// CFC twin of T_SafeMon_Tests: the same tests drawn as CFC diagrams, the way a TwinSAFE project is authored.
    FUNCTION_BLOCK T_SafeMon_Tests_CFC EXTENDS T_SafeCfcTestSuite
    VAR
    // Test_AutomaticRestartWhenGuardClosed
    group_1 : T_SafeGroup;
    fb_1 : T_SafeMon(group := group_1);
    // Test_SecureInputBypassesGuard
    group_2 : T_SafeGroup;
    fb_2 : T_SafeMon(group := group_2);
    // Test_ManualFunctionTestRequiresGuardOpenedOnce
    group_3 : T_SafeGroup;
    fb_3 : T_SafeMon(group := group_3) := (Parameters := (ManualFunctionTest := TRUE));
    // Test_EdmFaultWithoutManualRestartStaysSafe
    group_4 : T_SafeGroup;
    fb_4 : T_SafeMon(group := group_4);
END_VAR

Test_AutomaticRestartWhenGuardClosed();
Test_SecureInputBypassesGuard();
Test_ManualFunctionTestRequiresGuardOpenedOnce();
Test_EdmFaultWithoutManualRestartStaysSafe();

METHOD PRIVATE Test_AutomaticRestartWhenGuardClosed
// note: this text did not pass the execution check against the stored diagram
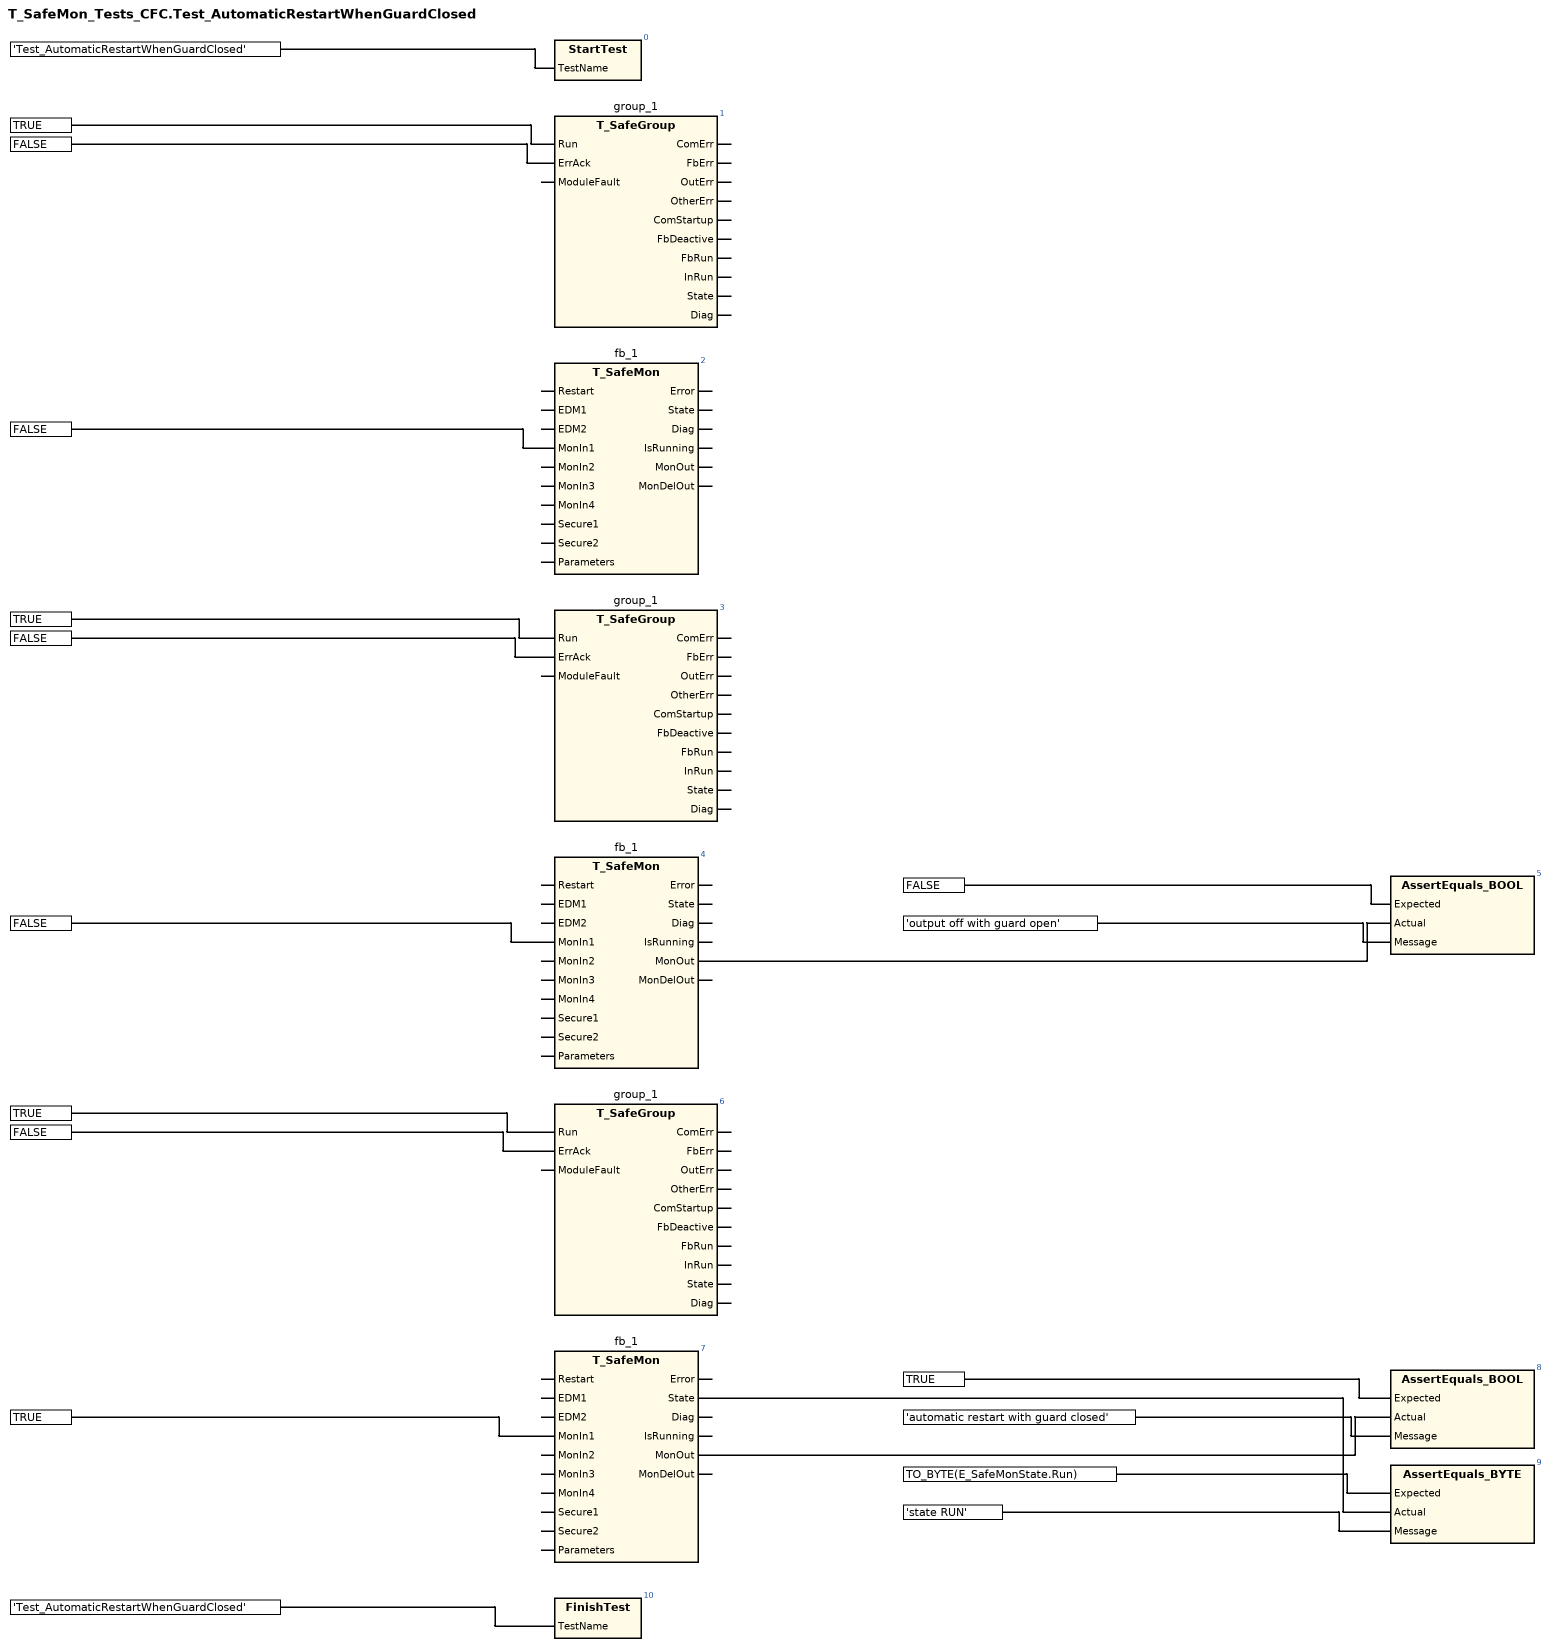
StartTest(TestName := 'Test_AutomaticRestartWhenGuardClosed');
group_1(Run := TRUE, ErrAck := FALSE); // T_SafeGroup
fb_1(MonIn1 := FALSE); // T_SafeMon
group_1(Run := TRUE, ErrAck := FALSE); // T_SafeGroup
fb_1(MonIn1 := FALSE); // T_SafeMon
AssertEquals_BOOL(Expected := FALSE, Actual := fb_1.MonOut, Message := 'output off with guard open');
group_1(Run := TRUE, ErrAck := FALSE); // T_SafeGroup
fb_1(MonIn1 := TRUE); // T_SafeMon
AssertEquals_BOOL(Expected := TRUE, Actual := fb_1.MonOut, Message := 'automatic restart with guard closed');
AssertEquals_BYTE(Expected := TO_BYTE(E_SafeMonState.Run), Actual := fb_1.State, Message := 'state RUN');
FinishTest(TestName := 'Test_AutomaticRestartWhenGuardClosed');
END_METHOD

METHOD PRIVATE Test_SecureInputBypassesGuard
// note: this text did not pass the execution check against the stored diagram
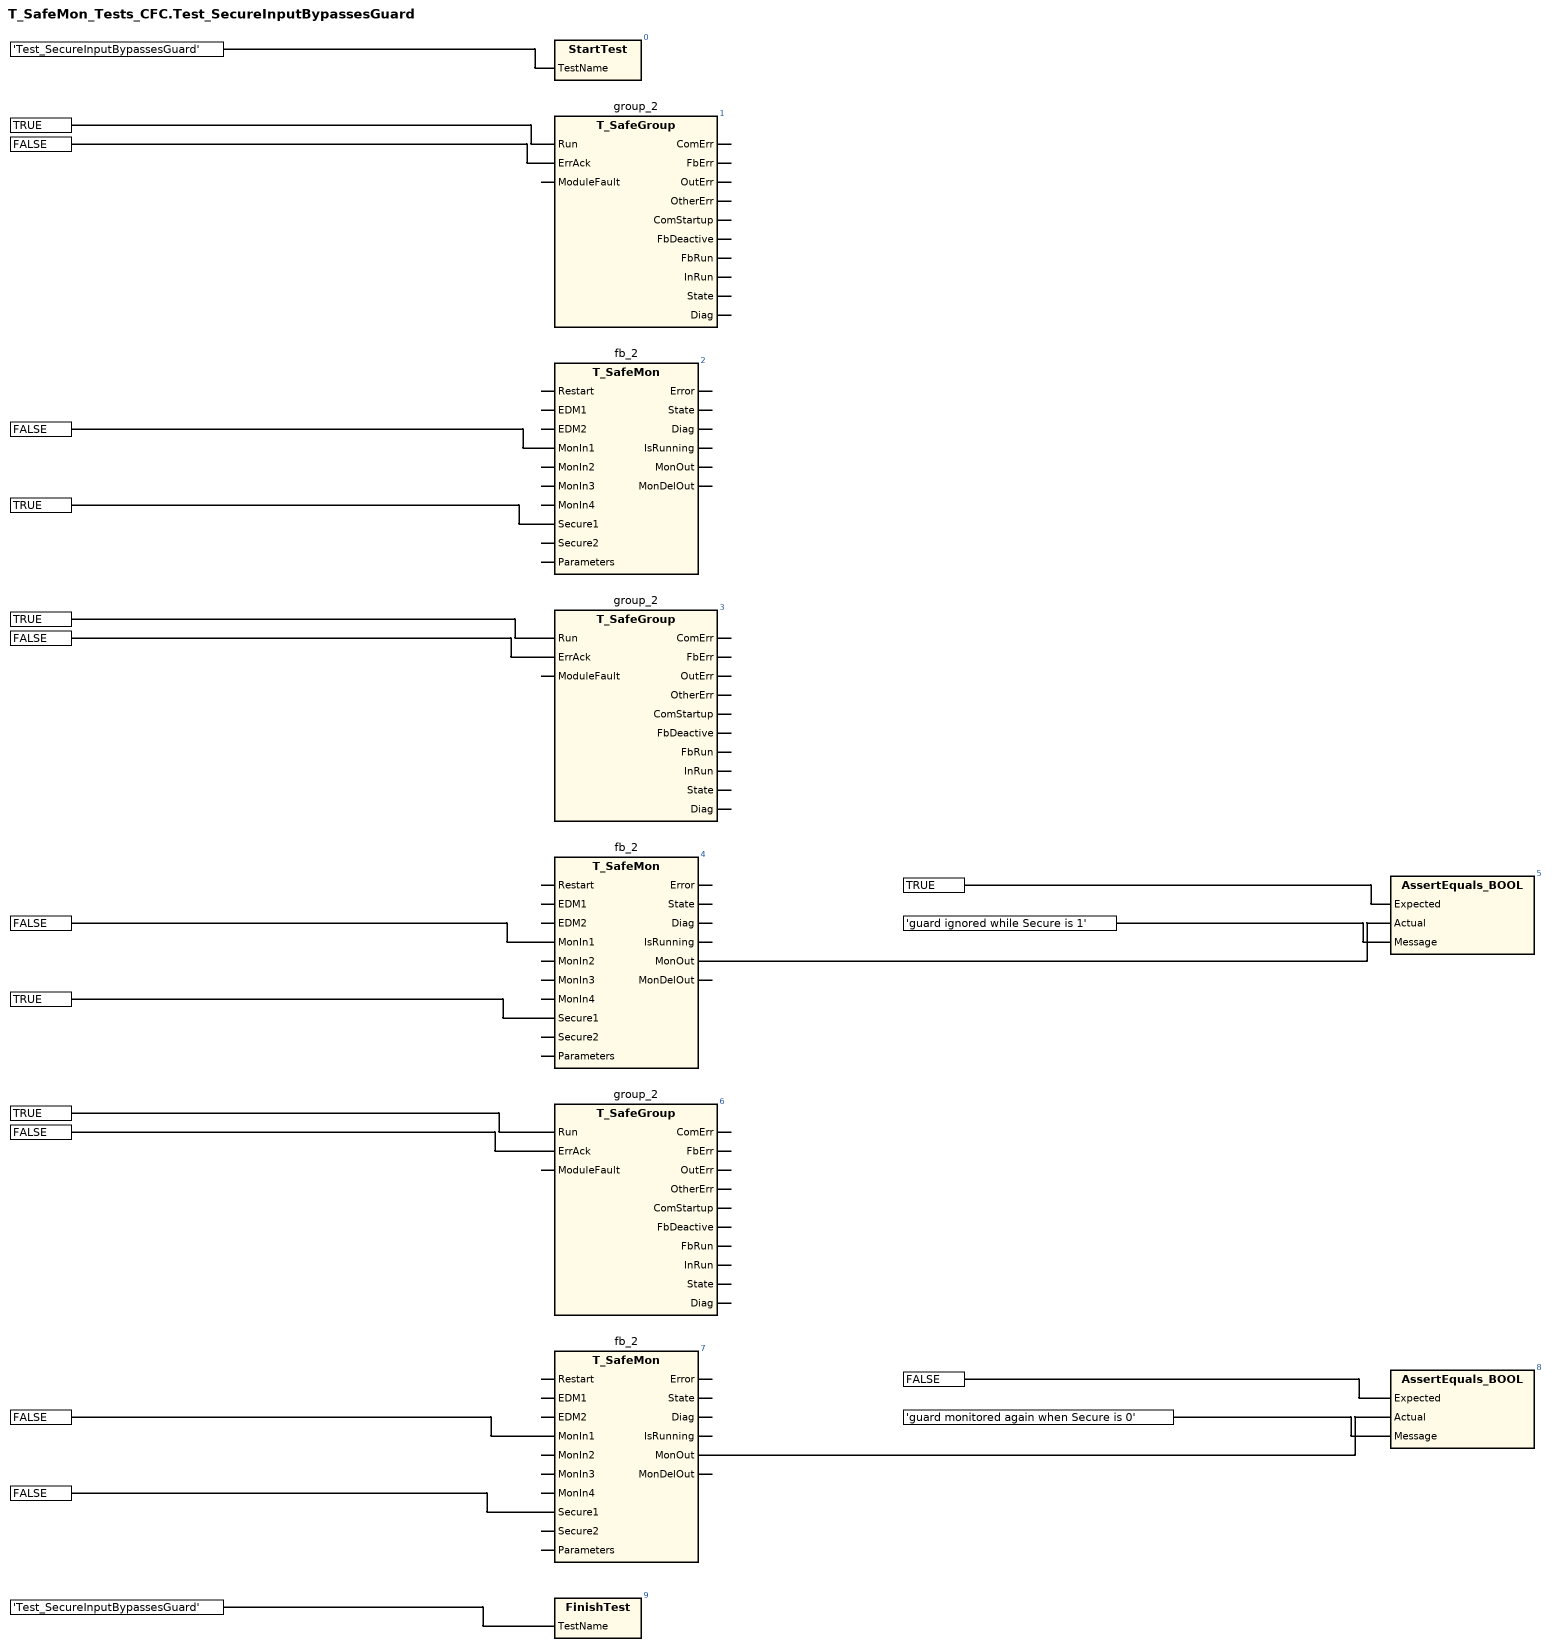
StartTest(TestName := 'Test_SecureInputBypassesGuard');
group_2(Run := TRUE, ErrAck := FALSE); // T_SafeGroup
fb_2(MonIn1 := FALSE, Secure1 := TRUE); // T_SafeMon
group_2(Run := TRUE, ErrAck := FALSE); // T_SafeGroup
fb_2(MonIn1 := FALSE, Secure1 := TRUE); // T_SafeMon
AssertEquals_BOOL(Expected := TRUE, Actual := fb_2.MonOut, Message := 'guard ignored while Secure is 1');
group_2(Run := TRUE, ErrAck := FALSE); // T_SafeGroup
fb_2(MonIn1 := FALSE, Secure1 := FALSE); // T_SafeMon
AssertEquals_BOOL(Expected := FALSE, Actual := fb_2.MonOut, Message := 'guard monitored again when Secure is 0');
FinishTest(TestName := 'Test_SecureInputBypassesGuard');
END_METHOD

METHOD PRIVATE Test_ManualFunctionTestRequiresGuardOpenedOnce
// note: this text did not pass the execution check against the stored diagram
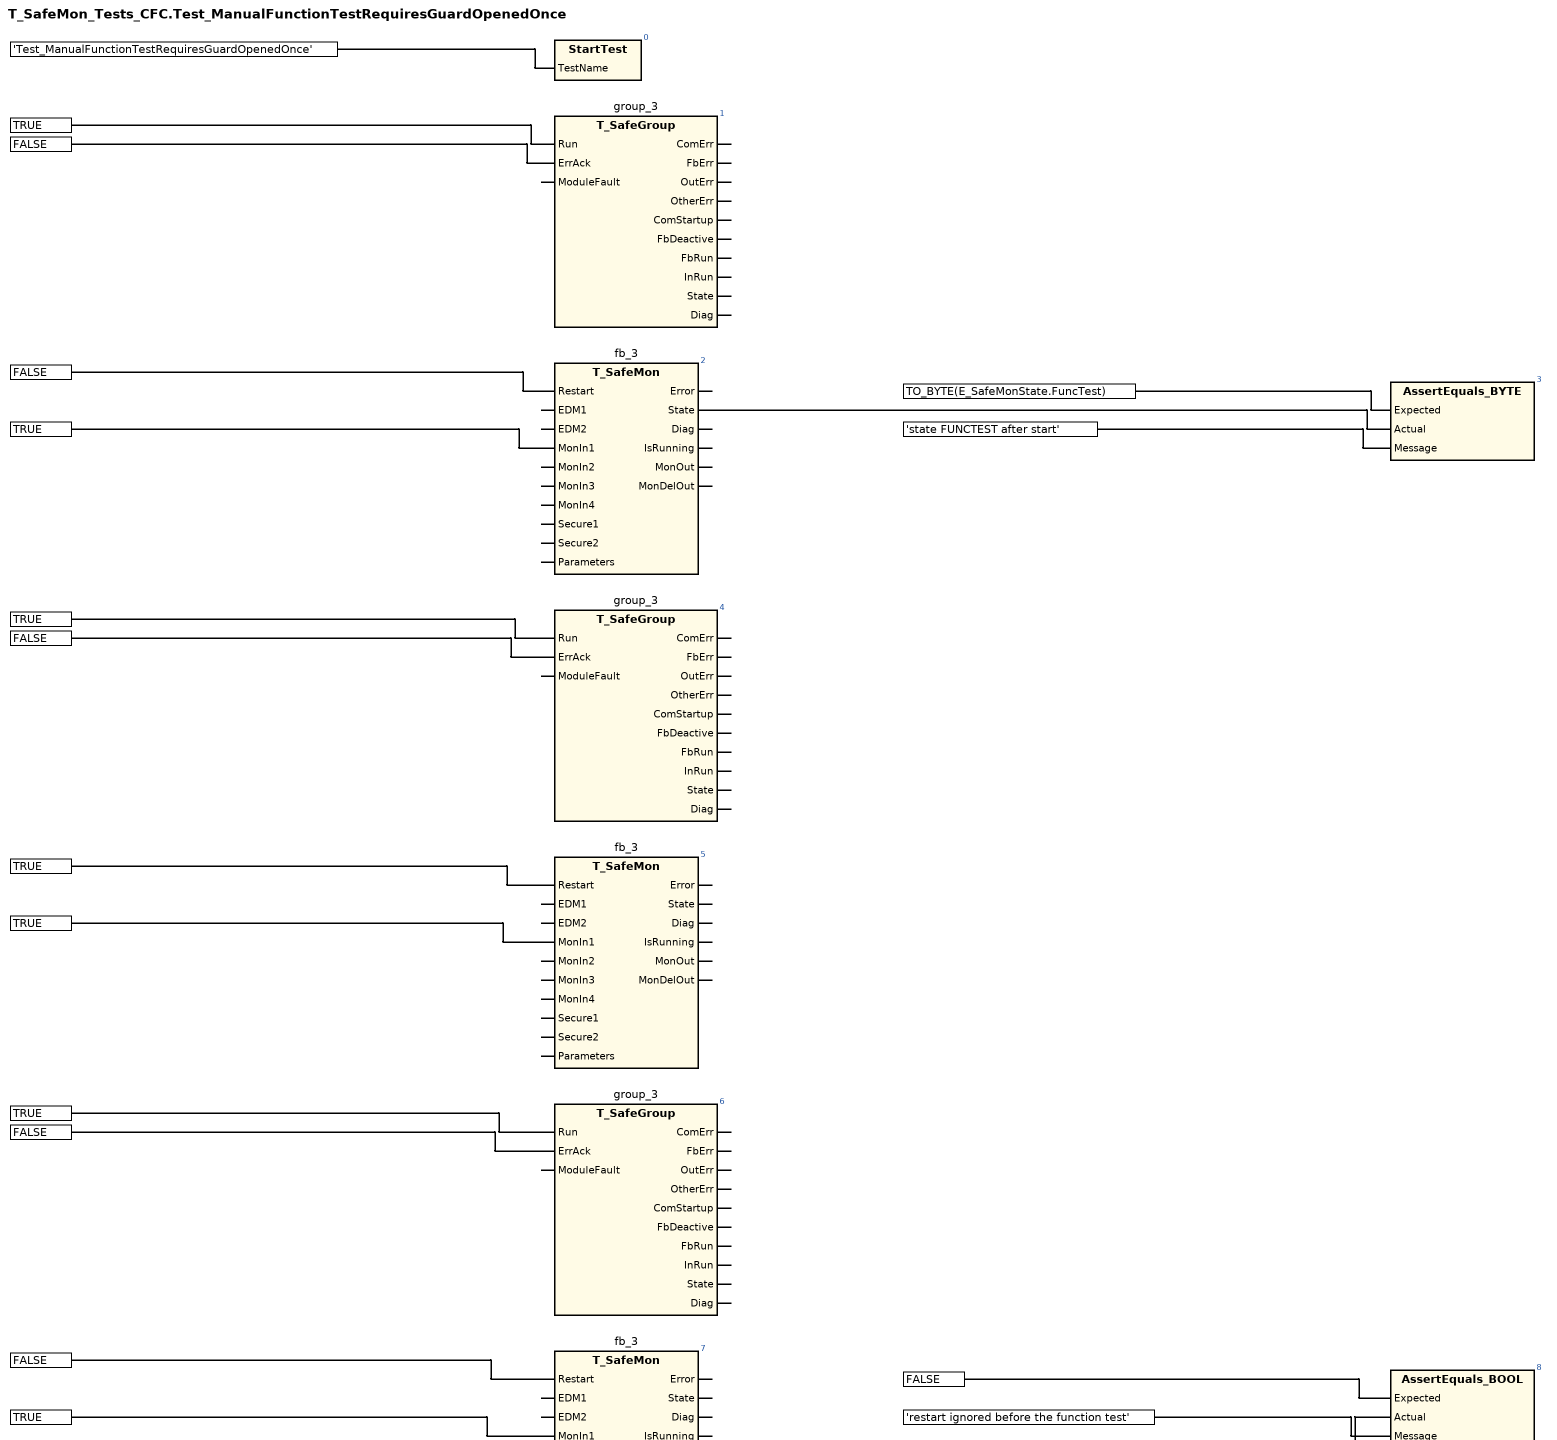
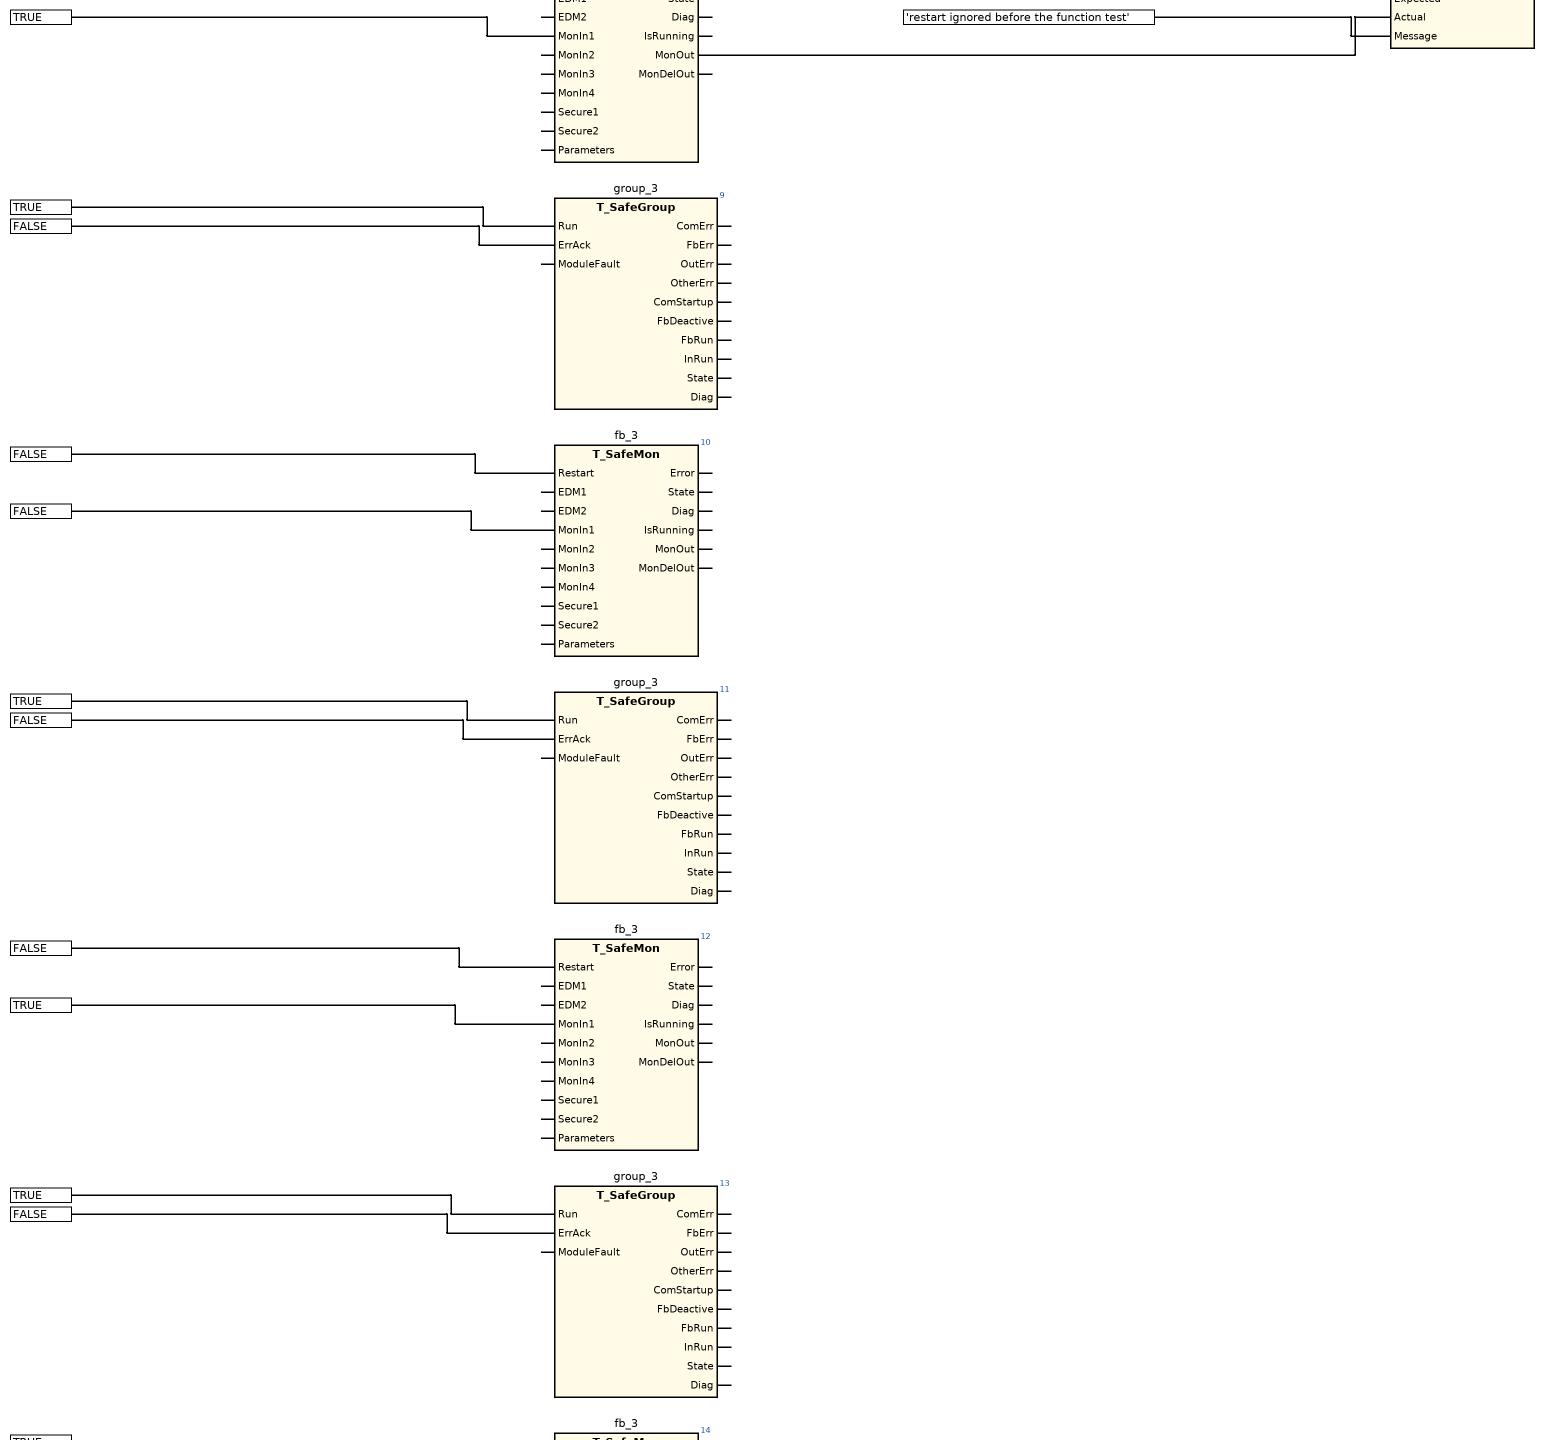
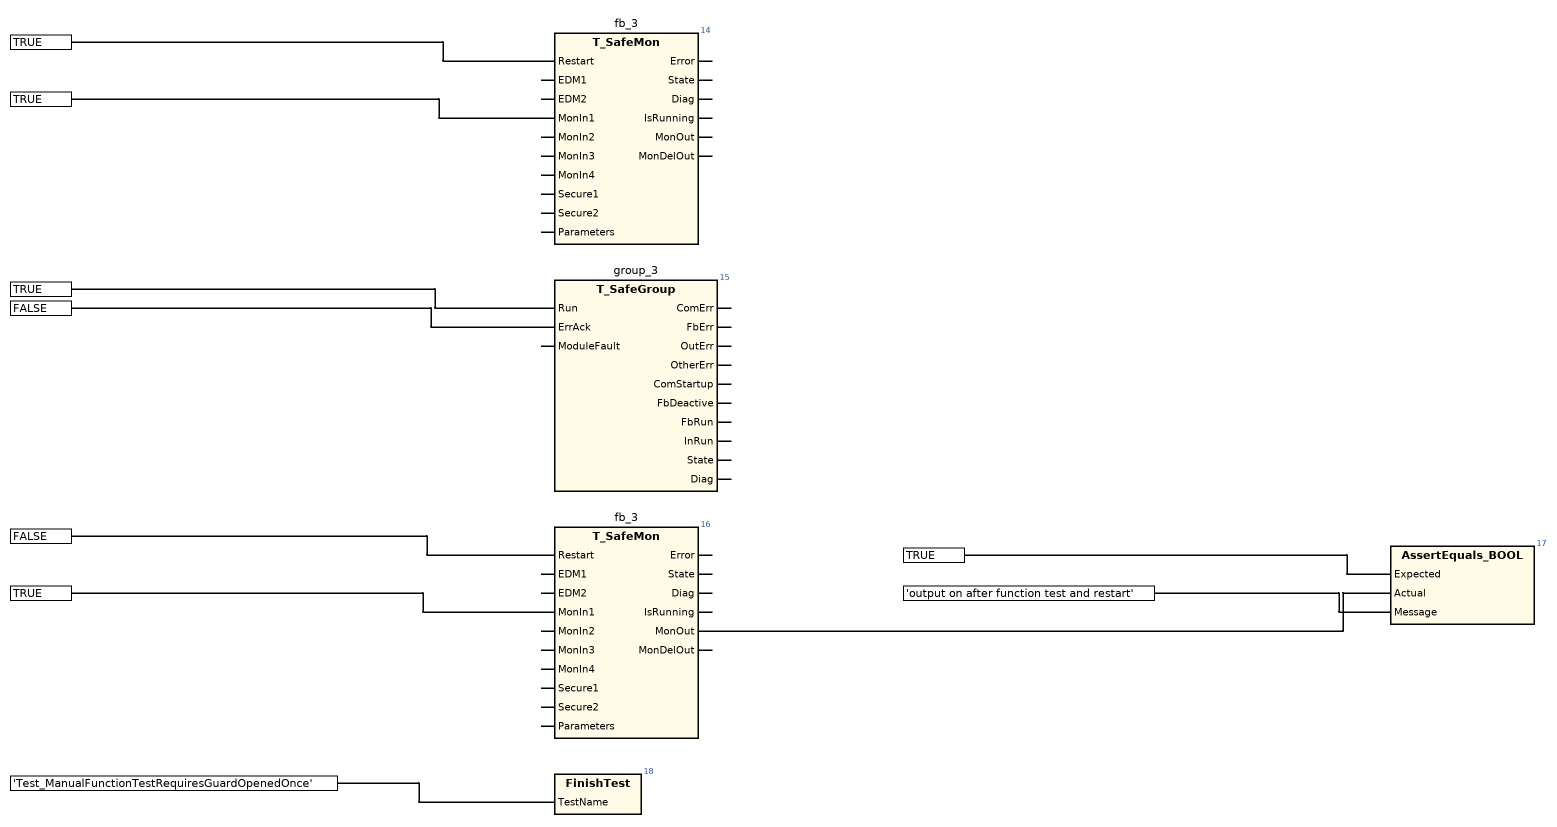
StartTest(TestName := 'Test_ManualFunctionTestRequiresGuardOpenedOnce');
group_3(Run := TRUE, ErrAck := FALSE); // T_SafeGroup
fb_3(Restart := FALSE, MonIn1 := TRUE); // T_SafeMon
AssertEquals_BYTE(Expected := TO_BYTE(E_SafeMonState.FuncTest), Actual := fb_3.State, Message := 'state FUNCTEST after start');
group_3(Run := TRUE, ErrAck := FALSE); // T_SafeGroup
fb_3(Restart := TRUE, MonIn1 := TRUE); // T_SafeMon
group_3(Run := TRUE, ErrAck := FALSE); // T_SafeGroup
fb_3(Restart := FALSE, MonIn1 := TRUE); // T_SafeMon
AssertEquals_BOOL(Expected := FALSE, Actual := fb_3.MonOut, Message := 'restart ignored before the function test');
group_3(Run := TRUE, ErrAck := FALSE); // T_SafeGroup
fb_3(Restart := FALSE, MonIn1 := FALSE); // T_SafeMon
group_3(Run := TRUE, ErrAck := FALSE); // T_SafeGroup
fb_3(Restart := FALSE, MonIn1 := TRUE); // T_SafeMon
group_3(Run := TRUE, ErrAck := FALSE); // T_SafeGroup
fb_3(Restart := TRUE, MonIn1 := TRUE); // T_SafeMon
group_3(Run := TRUE, ErrAck := FALSE); // T_SafeGroup
fb_3(Restart := FALSE, MonIn1 := TRUE); // T_SafeMon
AssertEquals_BOOL(Expected := TRUE, Actual := fb_3.MonOut, Message := 'output on after function test and restart');
FinishTest(TestName := 'Test_ManualFunctionTestRequiresGuardOpenedOnce');
END_METHOD

METHOD PRIVATE Test_EdmFaultWithoutManualRestartStaysSafe
// note: this text did not pass the execution check against the stored diagram
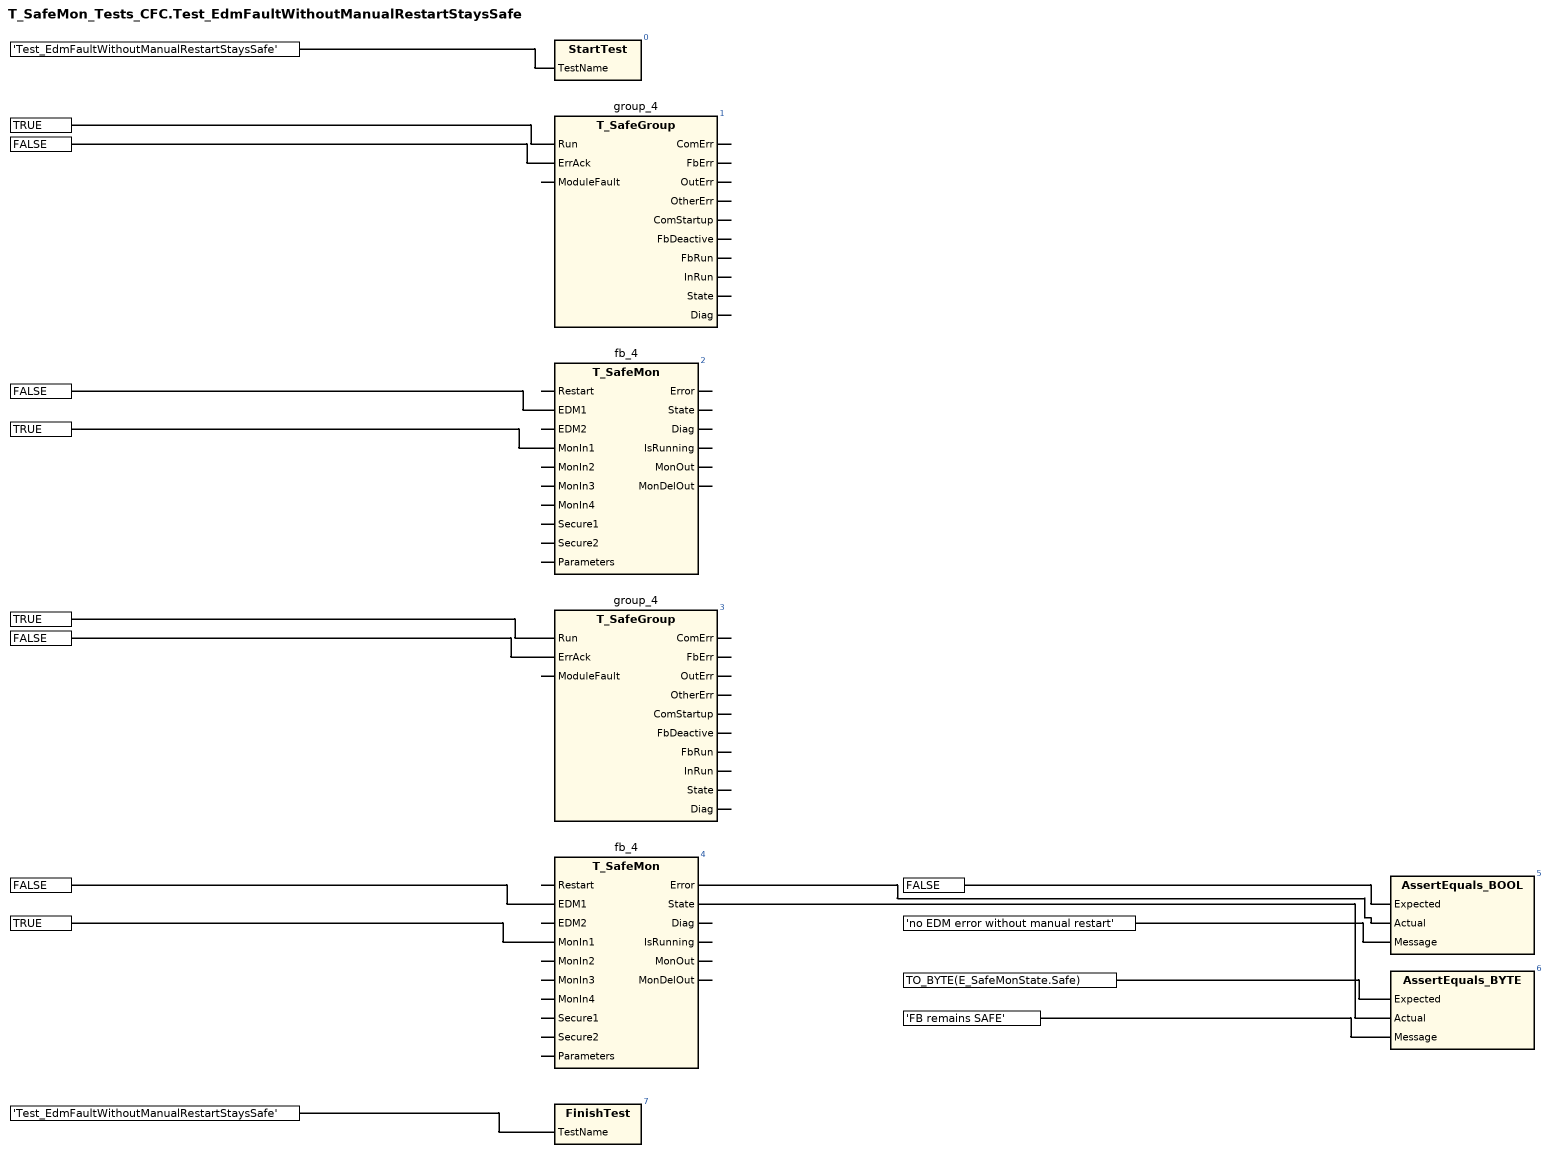
StartTest(TestName := 'Test_EdmFaultWithoutManualRestartStaysSafe');
group_4(Run := TRUE, ErrAck := FALSE); // T_SafeGroup
fb_4(EDM1 := FALSE, MonIn1 := TRUE); // T_SafeMon
group_4(Run := TRUE, ErrAck := FALSE); // T_SafeGroup
fb_4(EDM1 := FALSE, MonIn1 := TRUE); // T_SafeMon
AssertEquals_BOOL(Expected := FALSE, Actual := fb_4.Error, Message := 'no EDM error without manual restart');
AssertEquals_BYTE(Expected := TO_BYTE(E_SafeMonState.Safe), Actual := fb_4.State, Message := 'FB remains SAFE');
FinishTest(TestName := 'Test_EdmFaultWithoutManualRestartStaysSafe');
END_METHOD

END_FUNCTION_BLOCK

(* stored: Version 1.1.0.1, ProductVersion 3.1.4026.22
   POU T_SafeMon_Tests_CFC: Id {1d89c49f-59ee-5dfb-afa3-1bcdb112e803}, SpecialFunc None
   Method Test_AutomaticRestartWhenGuardClosed: Id {83b0d0c7-1361-574a-99ef-72935dbc2288}
   Method Test_SecureInputBypassesGuard: Id {a131705d-c025-589f-aeee-416054326699}
   Method Test_ManualFunctionTestRequiresGuardOpenedOnce: Id {d8f59f3e-7cf1-551d-8d89-88fbe46a68c4}
   Method Test_EdmFaultWithoutManualRestartStaysSafe: Id {67db55e4-cc93-5c85-976f-873a8e09b394} *)
